(* CODESYS project BODAS-RC18-12_27-18_40-DST.library
   Company: Bosch Rexroth AG
   DefaultNamespace: BODAS-RC18-12_27-18_40-DST
   Version: 2.3.0
   DocFormat: reStructuredText
   Description: User library to use BODAS-BDL services (API) for RC40.
   Title: BODAS_RC18-12_27-18_40-DST

Project tree, tasks and I/O mapping:
  DST/
    API/
      function bds_snsrDst_cfgSpdAndDir [ST]
      function bds_snsrDst_getSpdAndDir [ST]
      function bds_snsrDst_getTemp [ST]
    ENUM/
      data type bds_snsrDst_status_te
      data type bds_snsrDst_dir_te
    STRUCT/
      data type bds_snsrDst_cfgSpdAndDir_ts
      data type bds_snsrDst_statusDiag_tb
      data type bds_snsrDst_getSpdAndDir_ts
      data type bds_snsrDst_getTemp_ts
*)

// DST/ENUM/bds_snsrDst_status_te
{attribute 'external_name' := 'cmp_rts_bds_snsrDst_status_te'}
TYPE bds_snsrDst_status_te :
(
	bds_snsrDst_ok_E := 0,
	bds_snsrDst_outOfRange_E := 1,
	bds_snsrDst_frzn_E := 2,
	bds_snsrDst_standStill_E := 3,
	bds_snsrDst_err_E := 4,
	bds_snsrDst_invldConfig_E := 5,
	bds_snsrDst_notConfig_E := 6,
	bds_snsrDst_invldPrm_E := 7
)USINT;
END_TYPE

// DST/ENUM/bds_snsrDst_dir_te
{attribute 'external_name' := 'cmp_rts_bds_snsrDst_dir_te'}
TYPE bds_snsrDst_dir_te :
(
	bds_snsrDst_dirUnkown_E := 0,
	bds_snsrDst_dirClockwise_E := 1,
	bds_snsrDst_dirCounterClockwise_E := 2,
	bds_snsrDst_dirImpsChgErr_E := 3
)USINT;
END_TYPE

// DST/STRUCT/bds_snsrDst_cfgSpdAndDir_ts
{attribute 'external_name' := 'cmp_rts_bds_snsrDst_cfgSpdAndDir_ts'}
TYPE bds_snsrDst_cfgSpdAndDir_ts :
STRUCT 
	statusApi_e: bds_snsrDst_status_te; // statusApi_e 	        Status of the BDL function call
END_STRUCT
END_TYPE

// DST/STRUCT/bds_snsrDst_statusDiag_tb
(*Bit field type definition for the output module with diagnostic status information of output pin.*)
{attribute 'external_name' := 'cmp_rts_bds_snsrDst_statusDiag_tb'}
{attribute 'size' := '32'}
TYPE bds_snsrDst_statusDiag_tb :
STRUCT
	stErrSCB_b1: BIT; // Fault error status for short cut to battery
	stErrSCG_b1: BIT; // Fault error status for short cut to ground
	stErrOL_b1: BIT; // Fault error status for open load
	stErrOT_b1: BIT; // Fault error status for over temperature
	stErrUT_b1: BIT; // Fault error status for under temperature.
	stErrHw_b1: BIT; // Fault error status for hardware error for example  ADC connection is broken.
	resd1_b : ARRAY[0..2] OF BYTE;      (* Reserved *)
END_STRUCT
END_TYPE

// DST/STRUCT/bds_snsrDst_getSpdAndDir_ts
{attribute 'external_name' := 'cmp_rts_bds_snsrDst_getSpdAndDir_ts'}
TYPE bds_snsrDst_getSpdAndDir_ts :
STRUCT
	statusDiag_b: bds_snsrDst_statusDiag_tb; // statusDiag_b 	       Diagnostic information of sensor.
	spd_dRpm_u32: UDINT; // Rotation speed with resolution of 0.1 rpm.
	dir_e: bds_snsrDst_dir_te; // Rotation direction.
	statusApi_e: bds_snsrDst_status_te; // Status of the BDL API function call.
END_STRUCT
END_TYPE

// DST/STRUCT/bds_snsrDst_getTemp_ts
{attribute 'external_name' := 'cmp_rts_bds_snsrDst_getTemp_ts'}
TYPE bds_snsrDst_getTemp_ts :
STRUCT
	statusApi_e: bds_snsrDst_status_te; // Status of the BDL API function call.
	statusDiag_b: bds_snsrDst_statusDiag_tb; // Diagnostic information of sensor.
	temp_degC_s32: DINT; // Temperature in degree of celsius.
END_STRUCT
END_TYPE

// DST/API/bds_snsrDst_cfgSpdAndDir
/// The bds_snsrDst_cfgSpdAndDir API function configures the number of encoder wheel teeth.
///  
///==================================================================		  			===================================================================================================
///Return value    								  									     Description
///==================================================================		  			===================================================================================================
/// bds_snsrDst_cfgSpdAndDir_ts																	The return structure containing the status of API function call.																	
///
///==================================================================		   			===================================================================================================
///
///=======
///Code Example:
///=======
///============================================================================
///
/// PROGRAM OsInitProc
///VAR
///
///    bds_snsrDst_cfgSpdAndDir_s : bds_snsrDst_cfgSpdAndDir_ts;
///	
///    bds_snsrDst_inst_e : bds_snsrDst_inst_te;
///	
///    nrOfTeeth_u16 : UINT := 75;
///	
///END_VAR
///
///bds_snsrDst_inst_e := bds_snsrDst_inst_te.DrvPumpSpeed_E;
///
///bds_snsrDst_cfgSpdAndDir_s := bds_snsrDst_cfgSpdAndDir(bds_snsrDst_inst_e, nrOfTeeth_u16);
///
///IF bds_snsrDst_ok_E = bds_snsrDst_cfgSpdAndDir_s.statusApi_e THEN
///
///    (* configuration of DST sensor instance is successful *)
///	
///ELSE
///
///    (* error handling *)
///	
///END_IF;
/// END_PROGRAM
///
///============================================================================
{attribute 'external_name' := 'cmp_rts_bds_snsrDst_cfgSpdAndDir'}
FUNCTION bds_snsrDst_cfgSpdAndDir : bds_snsrDst_cfgSpdAndDir_ts
VAR_INPUT
	///The DST sensor instance name.
	snsrDstInst_e: USINT;
	///The number of wheel teeth for a particular DST sensor instance.
	///The range of wheel teeth is from 0 to 1000.
	nrOfTeeth_u16: UINT;
END_VAR

END_FUNCTION

// DST/API/bds_snsrDst_getSpdAndDir
/// The bds_snsrDst_getSpdAndDir API function provides calculated rotation speed with resolution of 0.1 rpm, rotation direction and diagnostic status of a particular DST sensor instance.
///
///Remarks
///
///A configuration function bds_snsrDst_cfgSpdAndDir is necessary, because calculation of rotation speed is based on number of wheel teeth.
///
///  
///==================================================================		  			===================================================================================================
///Return value    								  									     Description
///==================================================================		  			===================================================================================================
/// bds_snsrDst_getSpdAndDir_ts																	The return structure containing the status of API function call, wheel rotation speed in deci-rpm, wheel rotation direction and diagnostic information of a particular DST sensor instance. For detail information please refer into chapter DST.																
///
///==================================================================		   			===================================================================================================
///
///=======
///Code Example:
///=======
///============================================================================
///
/// PROGRAM OsInitProc
///VAR
///
///    bds_snsrDst_getSpdAndDir_s : bds_snsrDst_getSpdAndDir_ts;
///	
///    bds_snsrDst_inst_e : bds_snsrDst_inst_te;
///	
///    spd_dRpm_u32 : UDINT;
///	
///    rotDir_u8 : USINT;
///	
///END_VAR
///
///bds_snsrDst_inst_e := bds_snsrDst_inst_te.DrvPumpSpeed_E;
///
///bds_snsrDst_getSpdAndDir_s := bds_snsrDst_getSpdAndDir(bds_snsrDst_inst_e);
///
///IF bds_snsrDst_ok_E = bds_snsrDst_getSpdAndDir_s.statusApi_e THEN
///
///    (* save the actual wheel speed and rotation direction *)
///	
///    spd_dRpm_u32 := bds_snsrDst_getSpdAndDir_s.spd_dRpm_u32;
///	
///    rotDir_u8 := bds_snsrDst_getSpdAndDir_s.dir_e;
///	
///ELSE
///
///    (* error handling *)
///	
///END_IF;
/// END_PROGRAM
///
///============================================================================
{attribute 'external_name' := 'cmp_rts_bds_snsrDst_getSpdAndDir'}
FUNCTION bds_snsrDst_getSpdAndDir : bds_snsrDst_getSpdAndDir_ts
VAR_INPUT
	///The DST sensor instance name.
	snsrDstInst_e: USINT;
END_VAR

END_FUNCTION

// DST/API/bds_snsrDst_getTemp
/// The bds_snsrDst_getTemp API function provides temperature in degree celsius and diagnostic status of a particular DST sensor instance.
///  
///==================================================================		  			===================================================================================================
///Return value    								  									     Description
///==================================================================		  			===================================================================================================
/// bds_snsrDst_getTemp_ts																	The return structure containing the status of API function call, temperature in degree celsius and diagnostic information of a particular DST sensor instance. For detail information please refer into chapter DST.																
///
///==================================================================		   			===================================================================================================
///
///=======
///Code Example:
///=======
///============================================================================
///
/// PROGRAM OsInitProc
///VAR
///
///    bds_snsrDst_getTemp_s : bds_snsrDst_getTemp_ts;
///	
///    bds_snsrDst_inst_e : bds_snsrDst_inst_te;
///	
///    temp_degC_s32 : DINT;
///	
///END_VAR
///
///bds_snsrDst_inst_e := bds_snsrDst_inst_te.DrvPumpSpeed_E;
///
///bds_snsrDst_getTemp_s := bds_snsrDst_getTemp(bds_snsrDst_inst_e);
///
///IF bds_snsrDst_ok_E = bds_snsrDst_getTemp_s.statusApi_e THEN
///
///    (* save the actual temperature in degree celsius *)
///	
///    temp_degC_s32 := bds_snsrDst_getTemp_s.temp_degC_s32;
///	
///ELSE
///
///    (* error handling *)
///	
///END_IF;
/// END_PROGRAM
///
///============================================================================
{attribute 'external_name' := 'cmp_rts_bds_snsrDst_getTemp'}
FUNCTION bds_snsrDst_getTemp : bds_snsrDst_getTemp_ts
VAR_INPUT
	///The DST sensor instance name.
	snsrDstInst_e: USINT;
END_VAR

END_FUNCTION
